Fanuc KAREL source: KA00178.KL

PROGRAM KA00178
%NOLOCKGROUP
VAR
  SRC: ARRAY[4] OF STRING[20]
  DST: ARRAY[4] OF VECTOR
BEGIN
  DST = SRC
END KA00178
